(* Logix 5000 project; controller PickNPlace_Reto_2_SCADA Emulate 5570 rev 32.11; software revision 32.00 *)

TASK MainTask (continuous, watchdog 500 ms) : MainProgram

MODULES
   Local : Emulate 5570 (ICP 2, rev 32.11)
END_MODULES

VAR_GLOBAL   (* controller tags *)
   ALM_CAJA_NO_LLEGA : BOOL;   // Alarma: banda de entrada ON sin caja durante ALM_PRE_CAJA_NO_LLEGA
   ALM_CAJA_PERDIDA : BOOL;   // Alarma: la pinza perdio la caja durante el traslado (E5/E6)
   ALM_EMERGENCIA : BOOL;   // Alarma: parada de emergencia
   ALM_PINZA_VACIA : BOOL;   // Alarma: el brazo bajo (E3, Z quieto) y no tomo ninguna caja durante ALM_PRE_PINZA_VACIA
   ALM_PRE_CAJA_NO_LLEGA : DINT := 20000;   // Preset alarma caja no llega [ms] (configurable desde SCADA)
   ALM_PRE_CAJA_PERDIDA : DINT := 300;   // Preset alarma caja perdida [ms] (configurable desde SCADA)
   ALM_PRE_PINZA_VACIA : DINT := 2000;   // Preset alarma pinza vacia [ms] (configurable desde SCADA)
   ALM_PRE_ROBOT_NO_DISP : DINT := 10000;   // Preset alarma robot no disponible [ms] (configurable desde SCADA)
   ALM_ROBOT_NO_DISP : BOOL;   // Alarma: lote completo y robot sin READY durante ALM_PRE_ROBOT_NO_DISP
   CNT_CAJAS : DINT;   // Cajas contadas en Item at exit (flanco de E7)
   CNT_PRESET : DINT := 5;   // Cajas por lote
   ESTOP_ACTIVA : BOOL;   // Emergencia activa = X(S2)
   PROC_RUNNING : BOOL;   // Planta en marcha (alguna etapa E1..E10)
   PROC_WAIT_ROBOT : BOOL;   // Planta en pausa esperando al robot (E10)
   ROBOT_BUSY : BOOL;   // Robot ejecutando la rutina (Node-RED copia desde RAPID)
   ROBOT_DONE : BOOL;   // Robot termino la rutina (Node-RED copia desde RAPID)
   ROBOT_ESTOP : BOOL;   // Paro del robot por emergencia = X(S2) (Node-RED la copia a RAPID)
   ROBOT_READY : BOOL;   // Robot disponible (Node-RED copia desde RAPID)
   ROBOT_START : BOOL;   // Orden de rutina al robot = X(R1) (Node-RED la copia a RAPID)
   SCADA_ALM_ACK : BOOL;   // SCADA: reconocer alarmas
   SCADA_RESET : BOOL;   // SCADA: pulso de Reset tras emergencia
   SCADA_RESET_CNT : BOOL;   // SCADA: reiniciar contador de cajas (solo en R0)
   SCADA_START : BOOL;   // SCADA: pulso de marcha (Node-RED, trigger)
   SCADA_STOP : BOOL;   // SCADA: pulso de parada operativa
   STOP_CMD : BOOL;   // Parada operativa activa = X(S1)
END_VAR

PROGRAM MainProgram   (* main routine MainRoutine *)
VAR
   CV_101_01 : BOOL;
   E0 : BOOL;
   E1 : BOOL;
   E10 : BOOL;   // G1: pausa del lote, escena quieta esperando al robot
   E2 : BOOL;
   E2_FLAG_DELAY : TIMER := (PRE := 200);
   E3 : BOOL;
   E3_FLAG_DELAY : TIMER := (PRE := 200);
   E4 : BOOL;
   E4_FLAG : BOOL;
   E4_FLAG_DELAY : TIMER := (PRE := 500);
   E5 : BOOL;
   E5_FLAG_DELAY : TIMER := (PRE := 200);
   E6 : BOOL;
   E6_FLAG_DELAY : TIMER := (PRE := 200);
   E7 : BOOL;
   E7_FLAG_DELAY : TIMER := (PRE := 200);
   E7_ONS : BOOL;   // Memoria de flanco para contar cajas en E7
   E8 : BOOL;
   E8_FLAG_DELAY : TIMER := (PRE := 200);
   E9 : BOOL;
   E9_FLAG_DELAY : TIMER := (PRE := 200);
   R0 : BOOL;   // G2: esperando lote completo
   R1 : BOOL;   // G2: orden START al robot
   R2 : BOOL;   // G2: retirar orden y reiniciar conteo
   S0 : BOOL;   // G0: operacion normal
   S1 : BOOL;   // G0: STOP, forzado G1 a E0
   S2 : BOOL;   // G0: emergencia, forzado G1 vacio
   S3 : BOOL;   // G0: rearme, forzado G1 a E0
   SN_CV_101_01 : BOOL;
   SN_CV_101_01_ZS_01 : BOOL;
   SN_CV_101_01_ZS_02 : BOOL;
   SN_CV_101_02 : BOOL;
   SN_DSP_101_01 : INT;   // Factory IO: display Counter (= CNT_CAJAS)
   SN_PP01_AXIS_X_MOVING : BOOL;
   SN_PP01_AXIS_Z_MOVING : BOOL;
   SN_PP01_GR01 : BOOL;
   SN_PP01_GR01_ZS_01 : BOOL;
   SN_PP01_HS_01_START : BOOL;
   SN_PP01_HS_02_STOP : BOOL := 1;   // Factory IO: boton Stop (NC: 1 = sin presionar)
   SN_PP01_HS_03_ESTOP : BOOL := 1;   // Factory IO: parada de emergencia (NC: 1 = sin presionar)
   SN_PP01_HS_04_RESET : BOOL;   // Factory IO: boton Reset
   SN_PP01_MTR_X : BOOL;
   SN_PP01_MTR_Z : BOOL;
   START : BOOL;
   T1 : BOOL;
   T10 : BOOL;   // G1: lote completo y Pick & Place en reposo
   T11 : BOOL;   // G1: conteo reiniciado por G2 (robot DONE)
   T2 : BOOL;
   T3 : BOOL;
   T4 : BOOL;
   T5 : BOOL;
   T6 : BOOL;
   T7 : BOOL;
   T8 : BOOL;
   T9 : BOOL;
   TMR_CAJA_NO_LLEGA : TIMER := (PRE := 20000);   // Temporizador alarma caja no llega
   TMR_CAJA_PERDIDA : TIMER := (PRE := 300);   // Temporizador alarma caja perdida
   TMR_PINZA_VACIA : TIMER := (PRE := 2000);   // Temporizador alarma pinza vacia
   TMR_ROBOT_NO_DISP : TIMER := (PRE := 10000);   // Temporizador alarma robot no disponible
   TR1 : BOOL;   // G2: lote completo, robot READY y no BUSY, sin emergencia
   TR2 : BOOL;   // G2: ROBOT_DONE
   TR3 : BOOL;   // G2: DONE apagado
   TS1 : BOOL;   // G0: STOP local o SCADA sin emergencia
   TS2 : BOOL;   // G0: STOP liberado
   TS3 : BOOL;   // G0: hongo de emergencia presionado
   TS4 : BOOL;   // G0: hongo liberado y Reset
   TS5 : BOOL;   // G0: Reset liberado
END_VAR

ROUTINE MainRoutine   (* ladder *)
// Llamado ordenado de los 3 GRAFCET (G0 seguridad, G1 planta, G2 lote/robot) que corren en paralelo.
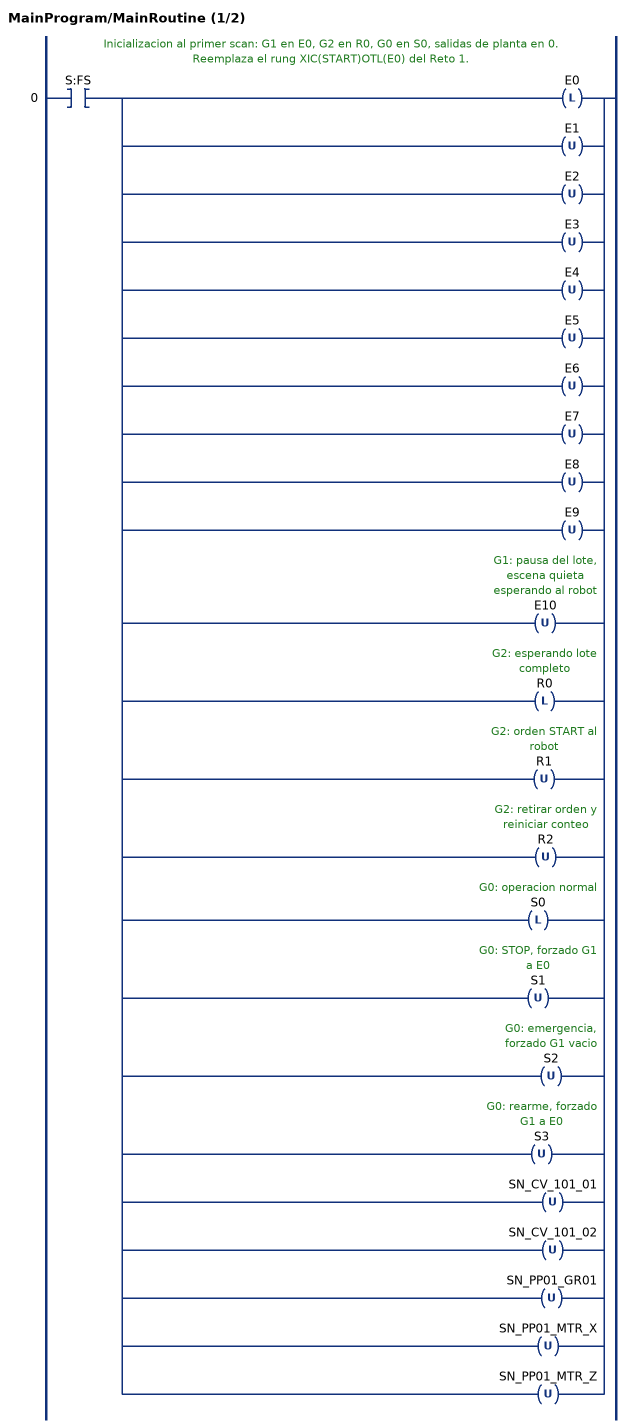
   // Inicializacion al primer scan: G1 en E0, G2 en R0, G0 en S0, salidas de planta en 0. Reemplaza el rung XIC(START)OTL(E0) del Reto 1.
   0: XIC(S:FS)[OTL(E0) ,OTU(E1) ,OTU(E2) ,OTU(E3) ,OTU(E4) ,OTU(E5) ,OTU(E6) ,OTU(E7) ,OTU(E8) ,OTU(E9) ,OTU(E10) ,OTL(R0) ,OTU(R1) ,OTU(R2) ,OTL(S0) ,OTU(S1) ,OTU(S2) ,OTU(S3) ,OTU(SN_CV_101_01) ,OTU(SN_CV_101_02) ,OTU(SN_PP01_GR01) ,OTU(SN_PP01_MTR_X) ,OTU(SN_PP01_MTR_Z) ];
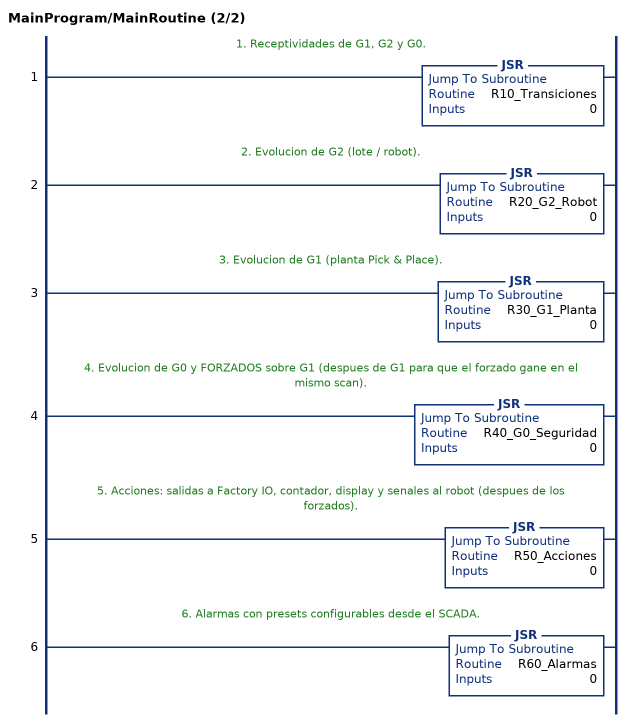
   // 1. Receptividades de G1, G2 y G0.
   1: JSR(R10_Transiciones,0);
   // 2. Evolucion de G2 (lote / robot).
   2: JSR(R20_G2_Robot,0);
   // 3. Evolucion de G1 (planta Pick & Place).
   3: JSR(R30_G1_Planta,0);
   // 4. Evolucion de G0 y FORZADOS sobre G1 (despues de G1 para que el forzado gane en el mismo scan).
   4: JSR(R40_G0_Seguridad,0);
   // 5. Acciones: salidas a Factory IO, contador, display y senales al robot (despues de los forzados).
   5: JSR(R50_Acciones,0);
   // 6. Alarmas con presets configurables desde el SCADA.
   6: JSR(R60_Alarmas,0);
END_ROUTINE

ROUTINE R10_Transiciones   (* ladder *)
// Receptividades (OTE) de los tres GRAFCET. T3..T9 son las del Reto 1 sin cambios.
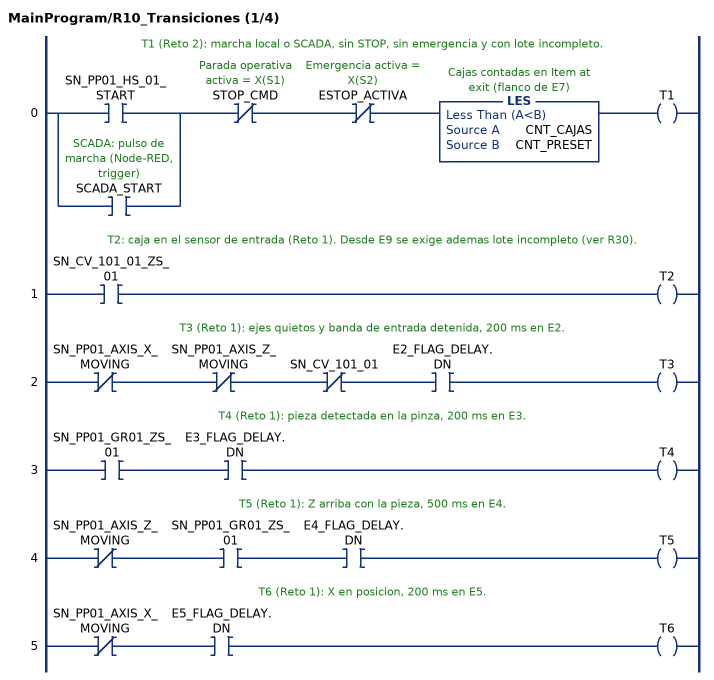
   // T1 (Reto 2): marcha local o SCADA, sin STOP, sin emergencia y con lote incompleto.
   0: [XIC(SN_PP01_HS_01_START) ,XIC(SCADA_START) ]XIO(STOP_CMD)XIO(ESTOP_ACTIVA)LES(CNT_CAJAS,CNT_PRESET)OTE(T1);
   // T2: caja en el sensor de entrada (Reto 1). Desde E9 se exige ademas lote incompleto (ver R30).
   1: XIC(SN_CV_101_01_ZS_01)OTE(T2);
   // T3 (Reto 1): ejes quietos y banda de entrada detenida, 200 ms en E2.
   2: XIO(SN_PP01_AXIS_X_MOVING)XIO(SN_PP01_AXIS_Z_MOVING)XIO(SN_CV_101_01)XIC(E2_FLAG_DELAY.DN)OTE(T3);
   // T4 (Reto 1): pieza detectada en la pinza, 200 ms en E3.
   3: XIC(SN_PP01_GR01_ZS_01)XIC(E3_FLAG_DELAY.DN)OTE(T4);
   // T5 (Reto 1): Z arriba con la pieza, 500 ms en E4.
   4: XIO(SN_PP01_AXIS_Z_MOVING)XIC(SN_PP01_GR01_ZS_01)XIC(E4_FLAG_DELAY.DN)OTE(T5);
   // T6 (Reto 1): X en posicion, 200 ms en E5.
   5: XIO(SN_PP01_AXIS_X_MOVING)XIC(E5_FLAG_DELAY.DN)OTE(T6);
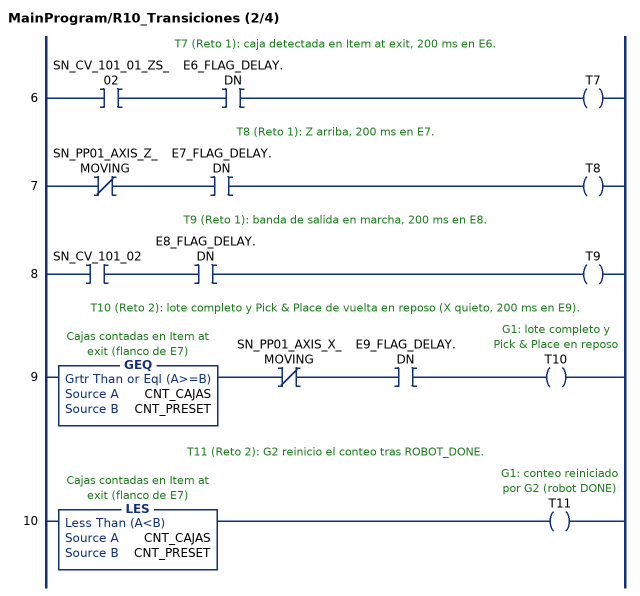
   // T7 (Reto 1): caja detectada en Item at exit, 200 ms en E6.
   6: XIC(SN_CV_101_01_ZS_02)XIC(E6_FLAG_DELAY.DN)OTE(T7);
   // T8 (Reto 1): Z arriba, 200 ms en E7.
   7: XIO(SN_PP01_AXIS_Z_MOVING)XIC(E7_FLAG_DELAY.DN)OTE(T8);
   // T9 (Reto 1): banda de salida en marcha, 200 ms en E8.
   8: XIC(SN_CV_101_02)XIC(E8_FLAG_DELAY.DN)OTE(T9);
   // T10 (Reto 2): lote completo y Pick & Place de vuelta en reposo (X quieto, 200 ms en E9).
   9: GEQ(CNT_CAJAS,CNT_PRESET)XIO(SN_PP01_AXIS_X_MOVING)XIC(E9_FLAG_DELAY.DN)OTE(T10);
   // T11 (Reto 2): G2 reinicio el conteo tras ROBOT_DONE.
   10: LES(CNT_CAJAS,CNT_PRESET)OTE(T11);
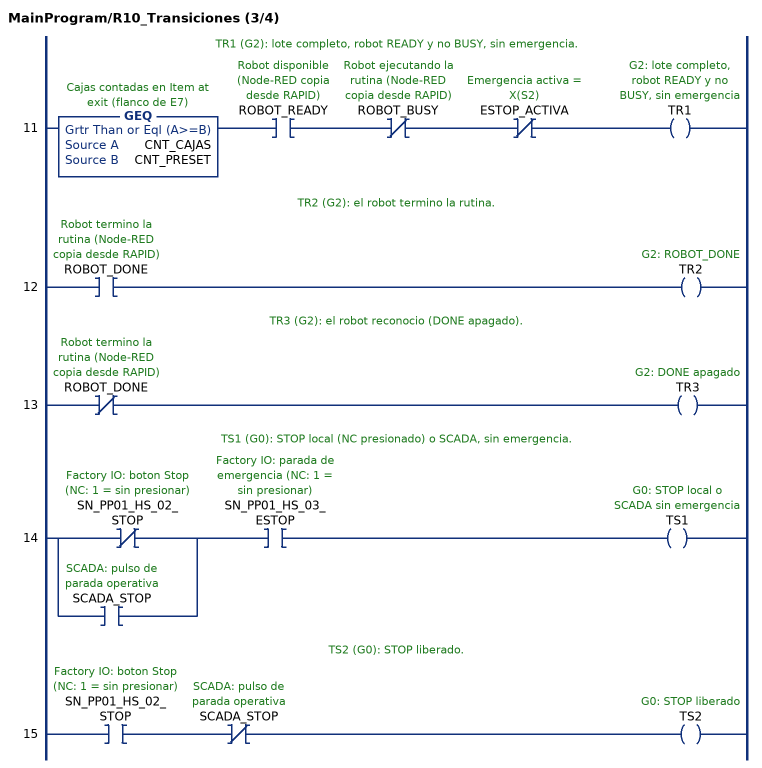
   // TR1 (G2): lote completo, robot READY y no BUSY, sin emergencia.
   11: GEQ(CNT_CAJAS,CNT_PRESET)XIC(ROBOT_READY)XIO(ROBOT_BUSY)XIO(ESTOP_ACTIVA)OTE(TR1);
   // TR2 (G2): el robot termino la rutina.
   12: XIC(ROBOT_DONE)OTE(TR2);
   // TR3 (G2): el robot reconocio (DONE apagado).
   13: XIO(ROBOT_DONE)OTE(TR3);
   // TS1 (G0): STOP local (NC presionado) o SCADA, sin emergencia.
   14: [XIO(SN_PP01_HS_02_STOP) ,XIC(SCADA_STOP) ]XIC(SN_PP01_HS_03_ESTOP)OTE(TS1);
   // TS2 (G0): STOP liberado.
   15: XIC(SN_PP01_HS_02_STOP)XIO(SCADA_STOP)OTE(TS2);
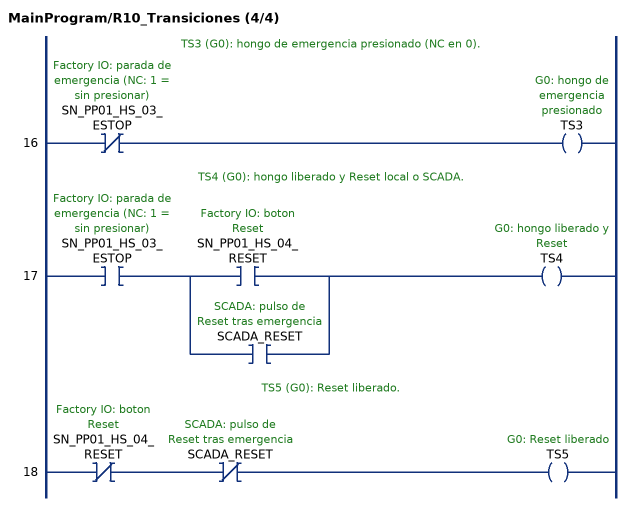
   // TS3 (G0): hongo de emergencia presionado (NC en 0).
   16: XIO(SN_PP01_HS_03_ESTOP)OTE(TS3);
   // TS4 (G0): hongo liberado y Reset local o SCADA.
   17: XIC(SN_PP01_HS_03_ESTOP)[XIC(SN_PP01_HS_04_RESET) ,XIC(SCADA_RESET) ]OTE(TS4);
   // TS5 (G0): Reset liberado.
   18: XIO(SN_PP01_HS_04_RESET)XIO(SCADA_RESET)OTE(TS5);
END_ROUTINE

ROUTINE R20_G2_Robot   (* ladder *)
// G2 Lote / robot: handshake READY / START / BUSY / DONE. No se fuerza con STOP.
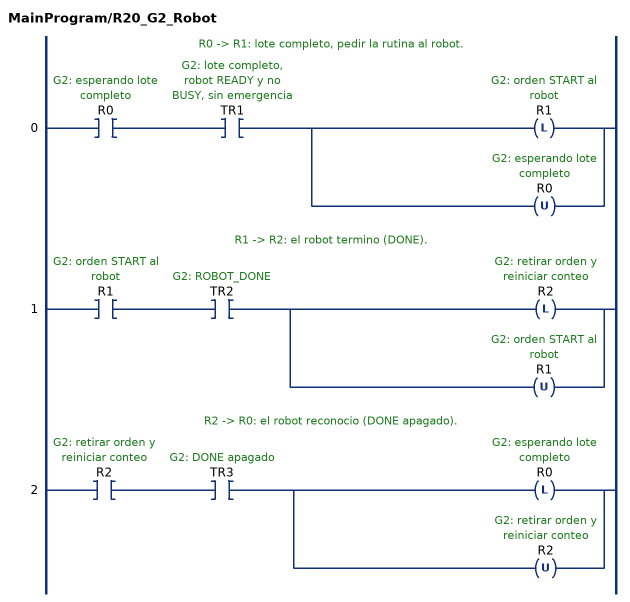
   // R0 -> R1: lote completo, pedir la rutina al robot.
   0: XIC(R0)XIC(TR1)[OTL(R1) ,OTU(R0) ];
   // R1 -> R2: el robot termino (DONE).
   1: XIC(R1)XIC(TR2)[OTL(R2) ,OTU(R1) ];
   // R2 -> R0: el robot reconocio (DONE apagado).
   2: XIC(R2)XIC(TR3)[OTL(R0) ,OTU(R2) ];
END_ROUTINE

ROUTINE R30_G1_Planta   (* ladder *)
// G1 Planta Pick & Place: GRAFCET del Reto 1 (E0..E9) + E10 (pausa del lote).
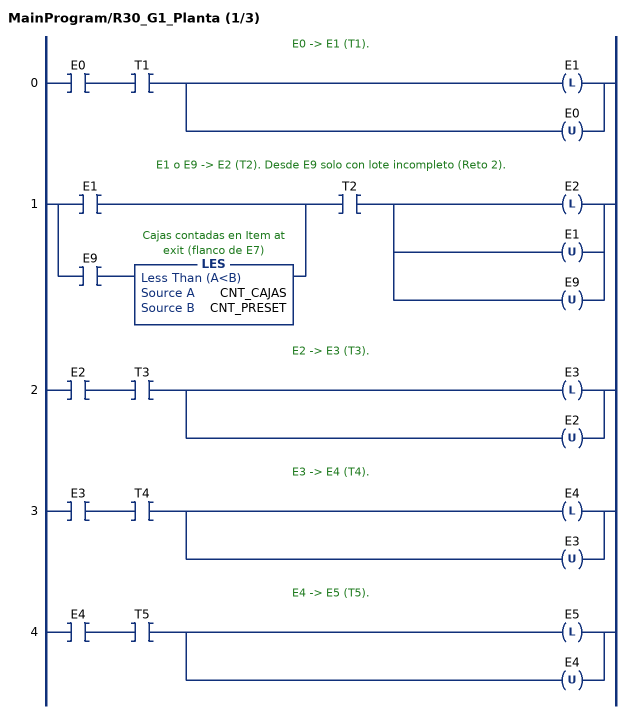
   // E0 -> E1 (T1).
   0: XIC(E0)XIC(T1)[OTL(E1) ,OTU(E0) ];
   // E1 o E9 -> E2 (T2). Desde E9 solo con lote incompleto (Reto 2).
   1: [XIC(E1) ,XIC(E9) LES(CNT_CAJAS,CNT_PRESET) ]XIC(T2)[OTL(E2) ,OTU(E1) ,OTU(E9) ];
   // E2 -> E3 (T3).
   2: XIC(E2)XIC(T3)[OTL(E3) ,OTU(E2) ];
   // E3 -> E4 (T4).
   3: XIC(E3)XIC(T4)[OTL(E4) ,OTU(E3) ];
   // E4 -> E5 (T5).
   4: XIC(E4)XIC(T5)[OTL(E5) ,OTU(E4) ];
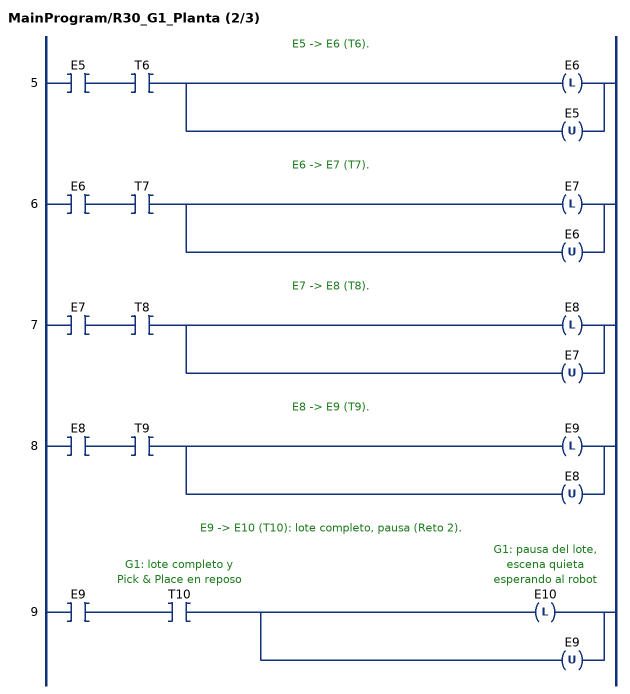
   // E5 -> E6 (T6).
   5: XIC(E5)XIC(T6)[OTL(E6) ,OTU(E5) ];
   // E6 -> E7 (T7).
   6: XIC(E6)XIC(T7)[OTL(E7) ,OTU(E6) ];
   // E7 -> E8 (T8).
   7: XIC(E7)XIC(T8)[OTL(E8) ,OTU(E7) ];
   // E8 -> E9 (T9).
   8: XIC(E8)XIC(T9)[OTL(E9) ,OTU(E8) ];
   // E9 -> E10 (T10): lote completo, pausa (Reto 2).
   9: XIC(E9)XIC(T10)[OTL(E10) ,OTU(E9) ];
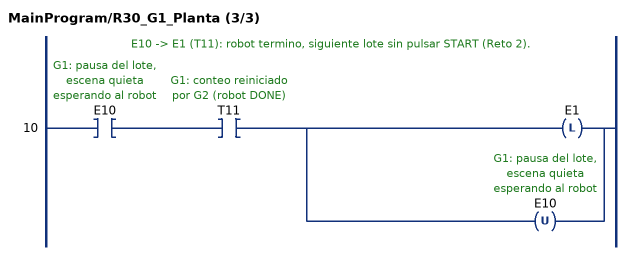
   // E10 -> E1 (T11): robot termino, siguiente lote sin pulsar START (Reto 2).
   10: XIC(E10)XIC(T11)[OTL(E1) ,OTU(E10) ];
END_ROUTINE

ROUTINE R40_G0_Seguridad   (* ladder *)
// G0 Seguridad y modos: STOP (forzado a E0) y emergencia (forzado vacio + Reset). Se ejecuta despues de G1.
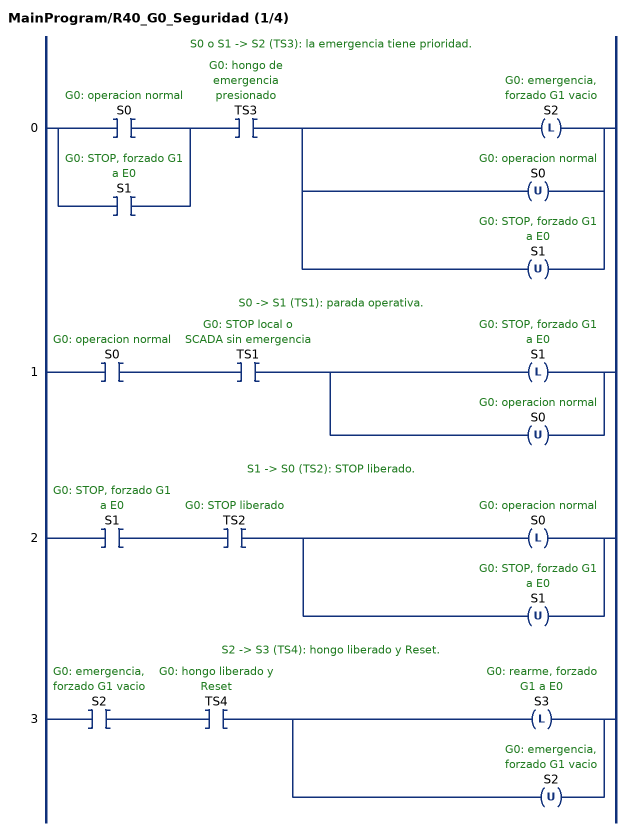
   // S0 o S1 -> S2 (TS3): la emergencia tiene prioridad.
   0: [XIC(S0) ,XIC(S1) ]XIC(TS3)[OTL(S2) ,OTU(S0) ,OTU(S1) ];
   // S0 -> S1 (TS1): parada operativa.
   1: XIC(S0)XIC(TS1)[OTL(S1) ,OTU(S0) ];
   // S1 -> S0 (TS2): STOP liberado.
   2: XIC(S1)XIC(TS2)[OTL(S0) ,OTU(S1) ];
   // S2 -> S3 (TS4): hongo liberado y Reset.
   3: XIC(S2)XIC(TS4)[OTL(S3) ,OTU(S2) ];
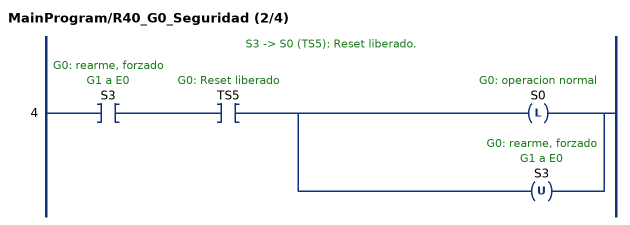
   // S3 -> S0 (TS5): Reset liberado.
   4: XIC(S3)XIC(TS5)[OTL(S0) ,OTU(S3) ];
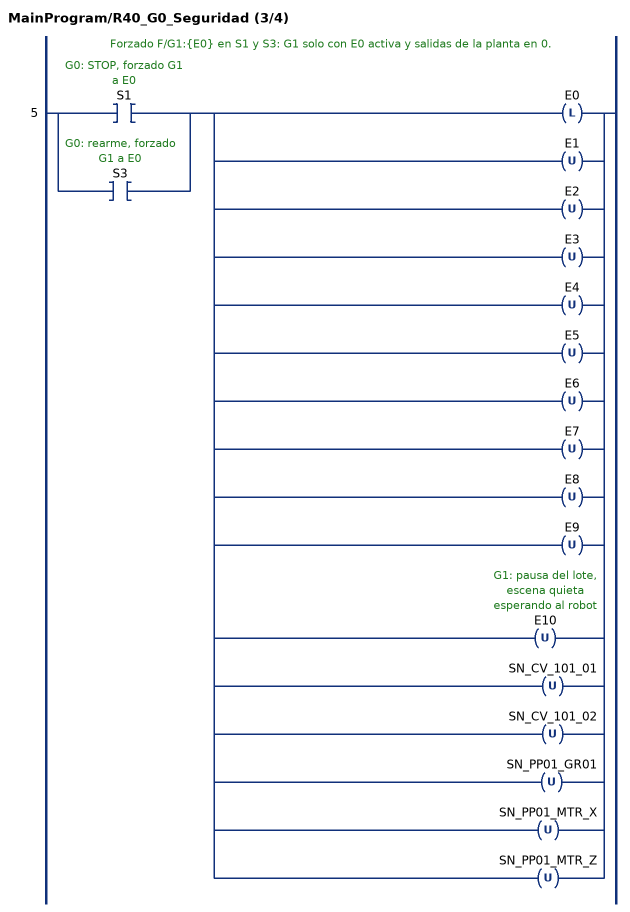
   // Forzado F/G1:{E0} en S1 y S3: G1 solo con E0 activa y salidas de la planta en 0.
   5: [XIC(S1) ,XIC(S3) ][OTL(E0) ,OTU(E1) ,OTU(E2) ,OTU(E3) ,OTU(E4) ,OTU(E5) ,OTU(E6) ,OTU(E7) ,OTU(E8) ,OTU(E9) ,OTU(E10) ,OTU(SN_CV_101_01) ,OTU(SN_CV_101_02) ,OTU(SN_PP01_GR01) ,OTU(SN_PP01_MTR_X) ,OTU(SN_PP01_MTR_Z) ];
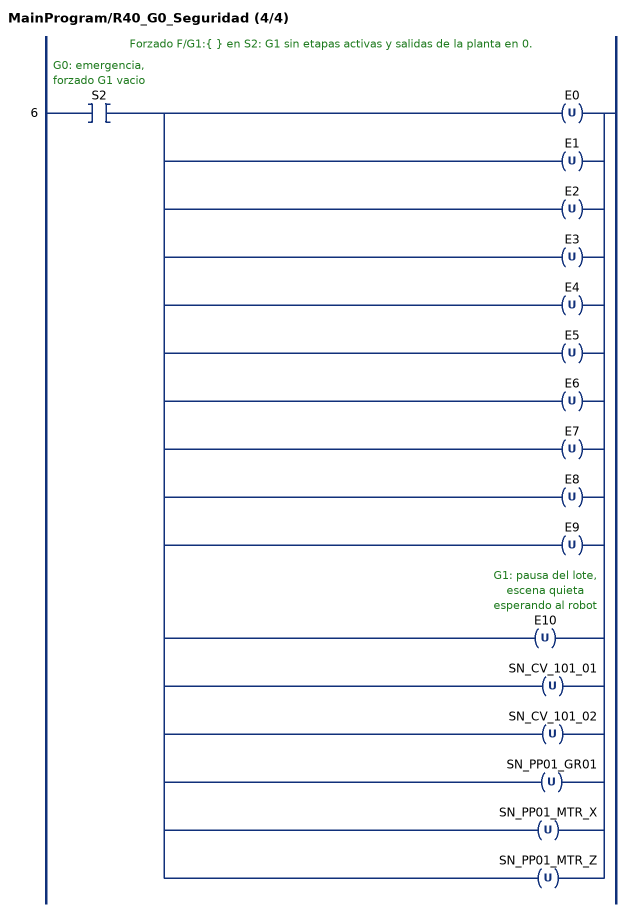
   // Forzado F/G1:{ } en S2: G1 sin etapas activas y salidas de la planta en 0.
   6: XIC(S2)[OTU(E0) ,OTU(E1) ,OTU(E2) ,OTU(E3) ,OTU(E4) ,OTU(E5) ,OTU(E6) ,OTU(E7) ,OTU(E8) ,OTU(E9) ,OTU(E10) ,OTU(SN_CV_101_01) ,OTU(SN_CV_101_02) ,OTU(SN_PP01_GR01) ,OTU(SN_PP01_MTR_X) ,OTU(SN_PP01_MTR_Z) ];
END_ROUTINE

ROUTINE R50_Acciones   (* ladder *)
// Acciones: las del Reto 1 sin cambios + E10, contador, display y senales a Node-RED.
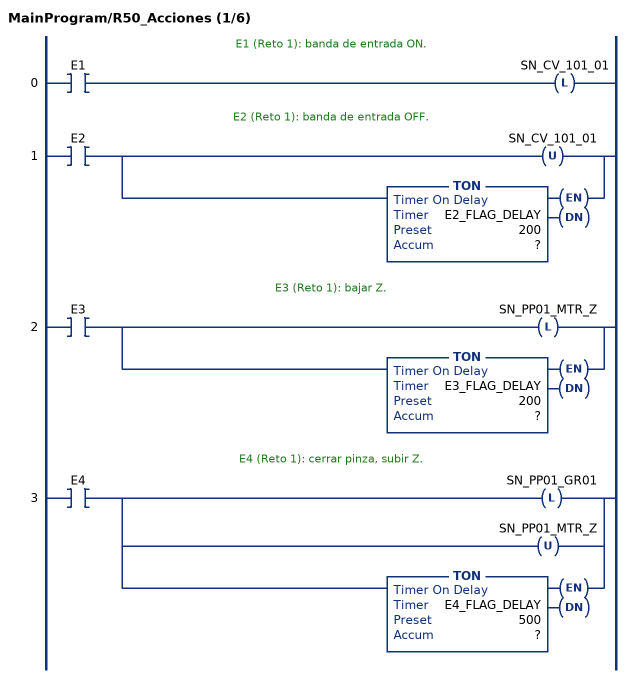
   // E1 (Reto 1): banda de entrada ON.
   0: XIC(E1)OTL(SN_CV_101_01);
   // E2 (Reto 1): banda de entrada OFF.
   1: XIC(E2)[OTU(SN_CV_101_01) ,TON(E2_FLAG_DELAY,?,?) ];
   // E3 (Reto 1): bajar Z.
   2: XIC(E3)[OTL(SN_PP01_MTR_Z) ,TON(E3_FLAG_DELAY,?,?) ];
   // E4 (Reto 1): cerrar pinza, subir Z.
   3: XIC(E4)[OTL(SN_PP01_GR01) ,OTU(SN_PP01_MTR_Z) ,TON(E4_FLAG_DELAY,?,?) ];
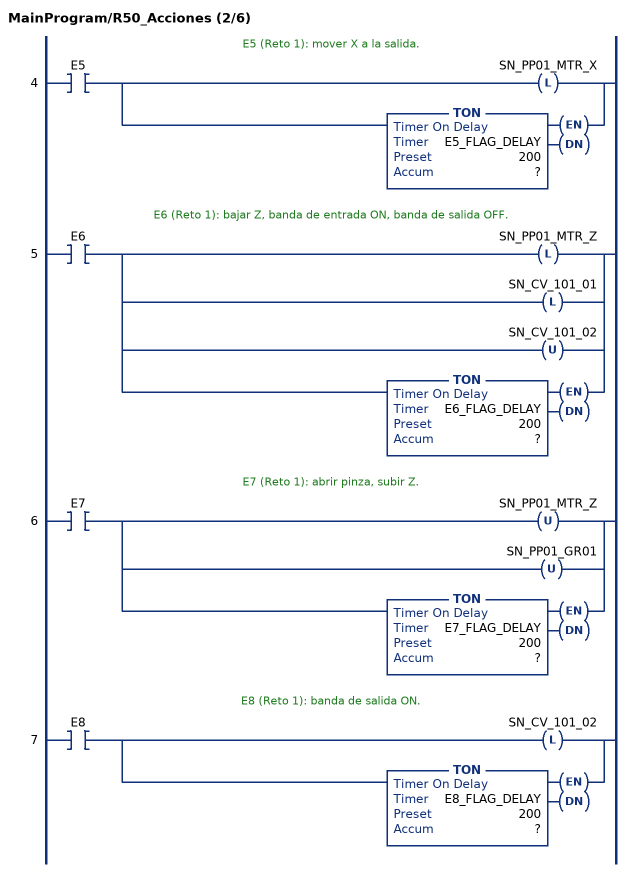
   // E5 (Reto 1): mover X a la salida.
   4: XIC(E5)[OTL(SN_PP01_MTR_X) ,TON(E5_FLAG_DELAY,?,?) ];
   // E6 (Reto 1): bajar Z, banda de entrada ON, banda de salida OFF.
   5: XIC(E6)[OTL(SN_PP01_MTR_Z) ,OTL(SN_CV_101_01) ,OTU(SN_CV_101_02) ,TON(E6_FLAG_DELAY,?,?) ];
   // E7 (Reto 1): abrir pinza, subir Z.
   6: XIC(E7)[OTU(SN_PP01_MTR_Z) ,OTU(SN_PP01_GR01) ,TON(E7_FLAG_DELAY,?,?) ];
   // E8 (Reto 1): banda de salida ON.
   7: XIC(E8)[OTL(SN_CV_101_02) ,TON(E8_FLAG_DELAY,?,?) ];
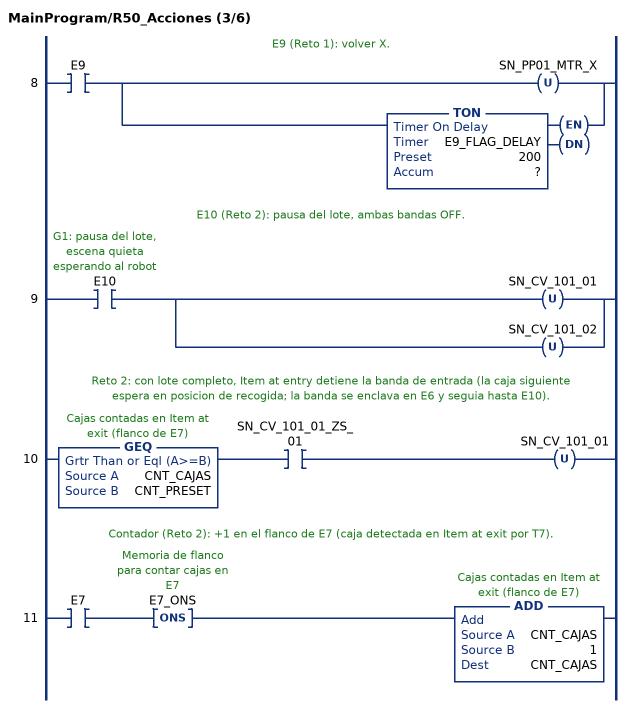
   // E9 (Reto 1): volver X.
   8: XIC(E9)[OTU(SN_PP01_MTR_X) ,TON(E9_FLAG_DELAY,?,?) ];
   // E10 (Reto 2): pausa del lote, ambas bandas OFF.
   9: XIC(E10)[OTU(SN_CV_101_01) ,OTU(SN_CV_101_02) ];
   // Reto 2: con lote completo, Item at entry detiene la banda de entrada (la caja siguiente espera en posicion de recogida; la banda se enclava en E6 y seguia hasta E10).
   10: GEQ(CNT_CAJAS,CNT_PRESET)XIC(SN_CV_101_01_ZS_01)OTU(SN_CV_101_01);
   // Contador (Reto 2): +1 en el flanco de E7 (caja detectada en Item at exit por T7).
   11: XIC(E7)ONS(E7_ONS)ADD(CNT_CAJAS,1,CNT_CAJAS);
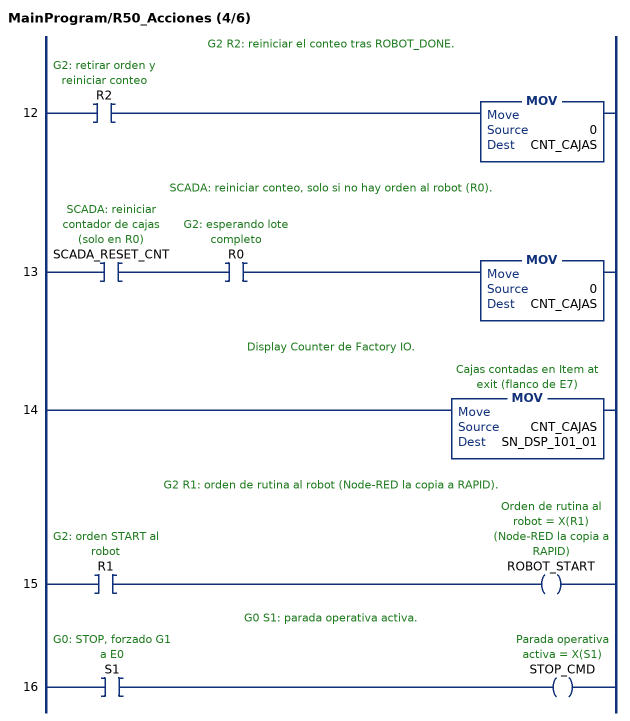
   // G2 R2: reiniciar el conteo tras ROBOT_DONE.
   12: XIC(R2)MOV(0,CNT_CAJAS);
   // SCADA: reiniciar conteo, solo si no hay orden al robot (R0).
   13: XIC(SCADA_RESET_CNT)XIC(R0)MOV(0,CNT_CAJAS);
   // Display Counter de Factory IO.
   14: MOV(CNT_CAJAS,SN_DSP_101_01);
   // G2 R1: orden de rutina al robot (Node-RED la copia a RAPID).
   15: XIC(R1)OTE(ROBOT_START);
   // G0 S1: parada operativa activa.
   16: XIC(S1)OTE(STOP_CMD);
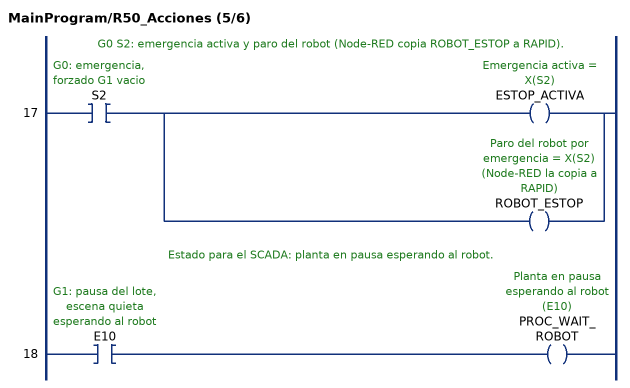
   // G0 S2: emergencia activa y paro del robot (Node-RED copia ROBOT_ESTOP a RAPID).
   17: XIC(S2)[OTE(ESTOP_ACTIVA) ,OTE(ROBOT_ESTOP) ];
   // Estado para el SCADA: planta en pausa esperando al robot.
   18: XIC(E10)OTE(PROC_WAIT_ROBOT);
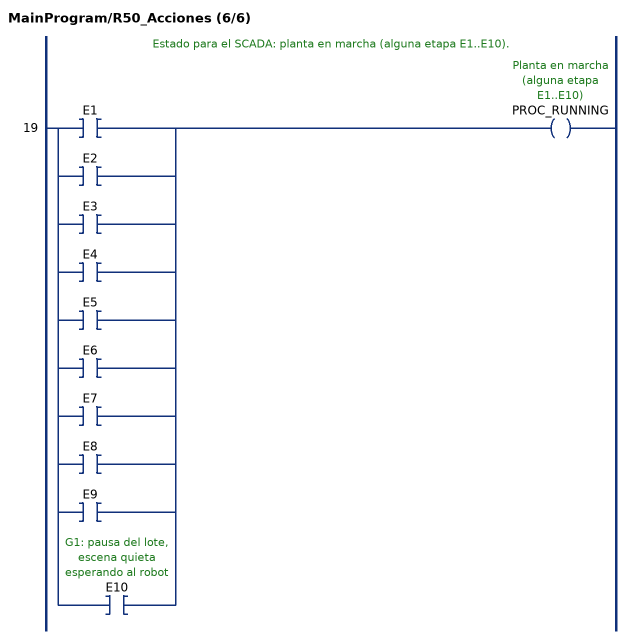
   // Estado para el SCADA: planta en marcha (alguna etapa E1..E10).
   19: [XIC(E1) ,XIC(E2) ,XIC(E3) ,XIC(E4) ,XIC(E5) ,XIC(E6) ,XIC(E7) ,XIC(E8) ,XIC(E9) ,XIC(E10) ]OTE(PROC_RUNNING);
END_ROUTINE

ROUTINE R60_Alarmas   (* ladder *)
// Alarmas del PLC. Presets en ms configurables desde el SCADA (ALM_PRE_*). Enclavadas hasta reconocer.
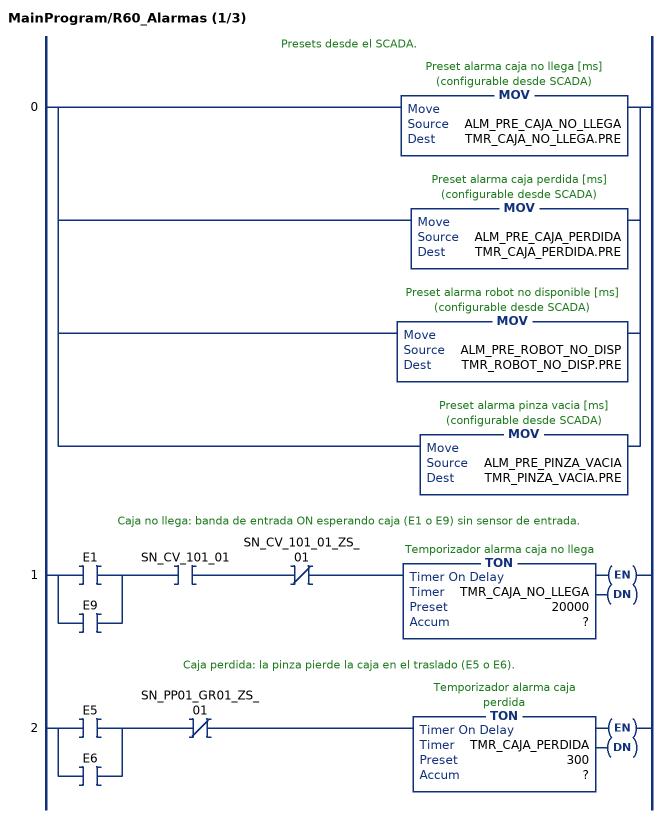
   // Presets desde el SCADA.
   0: [MOV(ALM_PRE_CAJA_NO_LLEGA,TMR_CAJA_NO_LLEGA.PRE) ,MOV(ALM_PRE_CAJA_PERDIDA,TMR_CAJA_PERDIDA.PRE) ,MOV(ALM_PRE_ROBOT_NO_DISP,TMR_ROBOT_NO_DISP.PRE) ,MOV(ALM_PRE_PINZA_VACIA,TMR_PINZA_VACIA.PRE) ];
   // Caja no llega: banda de entrada ON esperando caja (E1 o E9) sin sensor de entrada.
   1: [XIC(E1) ,XIC(E9) ]XIC(SN_CV_101_01)XIO(SN_CV_101_01_ZS_01)TON(TMR_CAJA_NO_LLEGA,?,?);
   // Caja perdida: la pinza pierde la caja en el traslado (E5 o E6).
   2: [XIC(E5) ,XIC(E6) ]XIO(SN_PP01_GR01_ZS_01)TON(TMR_CAJA_PERDIDA,?,?);
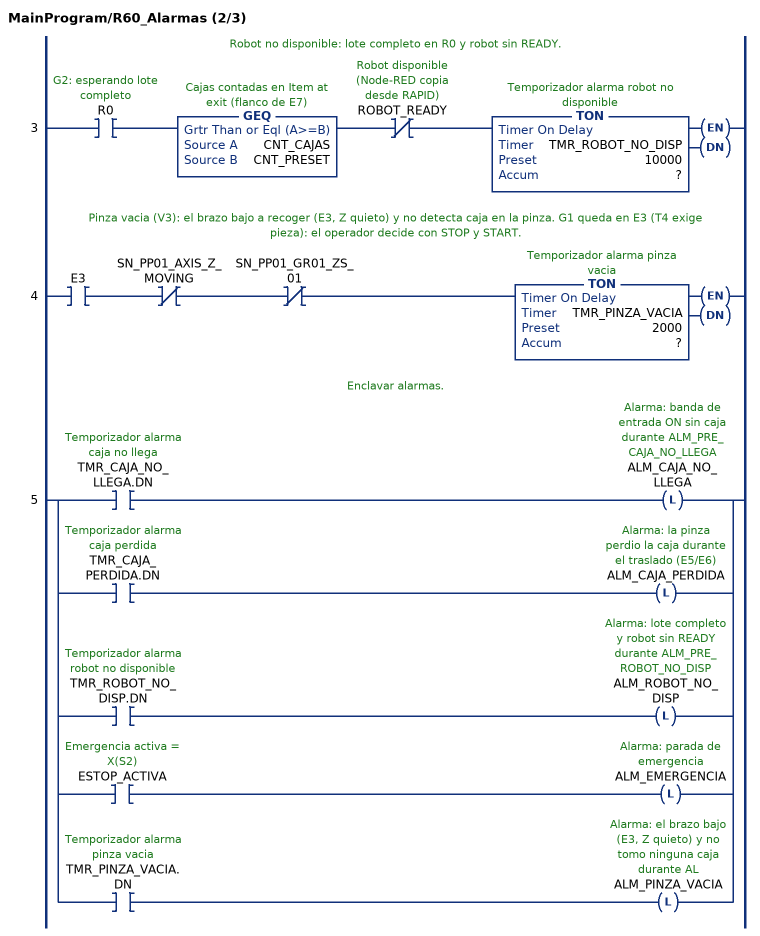
   // Robot no disponible: lote completo en R0 y robot sin READY.
   3: XIC(R0)GEQ(CNT_CAJAS,CNT_PRESET)XIO(ROBOT_READY)TON(TMR_ROBOT_NO_DISP,?,?);
   // Pinza vacia (V3): el brazo bajo a recoger (E3, Z quieto) y no detecta caja en la pinza. G1 queda en E3 (T4 exige pieza): el operador decide con STOP y START.
   4: XIC(E3)XIO(SN_PP01_AXIS_Z_MOVING)XIO(SN_PP01_GR01_ZS_01)TON(TMR_PINZA_VACIA,?,?);
   // Enclavar alarmas.
   5: [XIC(TMR_CAJA_NO_LLEGA.DN) OTL(ALM_CAJA_NO_LLEGA) ,XIC(TMR_CAJA_PERDIDA.DN) OTL(ALM_CAJA_PERDIDA) ,XIC(TMR_ROBOT_NO_DISP.DN) OTL(ALM_ROBOT_NO_DISP) ,XIC(ESTOP_ACTIVA) OTL(ALM_EMERGENCIA) ,XIC(TMR_PINZA_VACIA.DN) OTL(ALM_PINZA_VACIA) ];
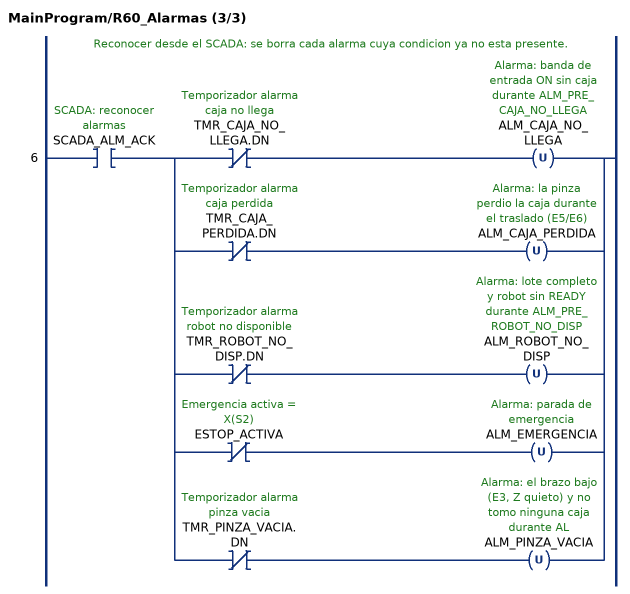
   // Reconocer desde el SCADA: se borra cada alarma cuya condicion ya no esta presente.
   6: XIC(SCADA_ALM_ACK)[XIO(TMR_CAJA_NO_LLEGA.DN) OTU(ALM_CAJA_NO_LLEGA) ,XIO(TMR_CAJA_PERDIDA.DN) OTU(ALM_CAJA_PERDIDA) ,XIO(TMR_ROBOT_NO_DISP.DN) OTU(ALM_ROBOT_NO_DISP) ,XIO(ESTOP_ACTIVA) OTU(ALM_EMERGENCIA) ,XIO(TMR_PINZA_VACIA.DN) OTU(ALM_PINZA_VACIA) ];
END_ROUTINE
END_PROGRAM
